(* LS Electric XG5000 project: GRST *)
(* PLC LSPLC *)

PROGRAM NewProgram (* task: 스캔 프로그램 *)
VAR
    Count : INT; (* Source preservation check *)
END_VAR
Count := Count + 1;
END_PROGRAM

PROGRAM AddedST (* task: 스캔 프로그램 *)
VAR
    Count : INT; (* Source preservation check *)
END_VAR
Count := Count + 1;
END_PROGRAM

PROGRAM AddedIL (* task: 스캔 프로그램 *)
VAR
    Count : INT; (* Source preservation check *)
END_VAR
LD Count
ADD 1
ST Count
END_PROGRAM